Fanuc KAREL source: KT00229.KL

PROGRAM KT00229
%NOLOCKGROUP
VAR
  B1: BOOLEAN
  Y2: ARRAY[2] OF BYTE
  OUT: BOOLEAN
BEGIN
  B1 = TRUE
    Y2[1] = 3
  OUT = B1 OR Y2[1]
END KT00229
